Fanuc KAREL source: KT00695.KL

PROGRAM KT00695
%NOLOCKGROUP
VAR
  V1: VECTOR
  V2: VECTOR
  OUT: REAL
BEGIN
  V1.X = 1.0
  V2.Y = 2.0
  V1.X = 1.0
  V2.Y = 2.0
  OUT = - V1
END KT00695
